(* Logix 5000 project; controller R400_500_XLS vendor 1 type 14 code 216 rev 31.11; software revision 31.01; part 32 of 32 *)
(* tags used below, declared in another part *)
   CycExcBuffer : UDT_CYCLE;
   CycleSequence : UDT_CYCLE_SEQUENCE;
   DRYING : DINT;   // Drying id number
   FINALRINSE_1 : DINT;   // Final rinse 1 id number
   M : DINT[5];   // Memory Bits
   OneShot : DINT[1];
   RINSE_4 : DINT;   // Rinse 4 id number
   RinseExcBuffer : UDT_RINSE;
   VENTING : DINT;   // Venting id number
   TreatmentPtr : DINT;
   Unit : Hrdwre;   // Unit Configuration
(* MainProgram, continued *)

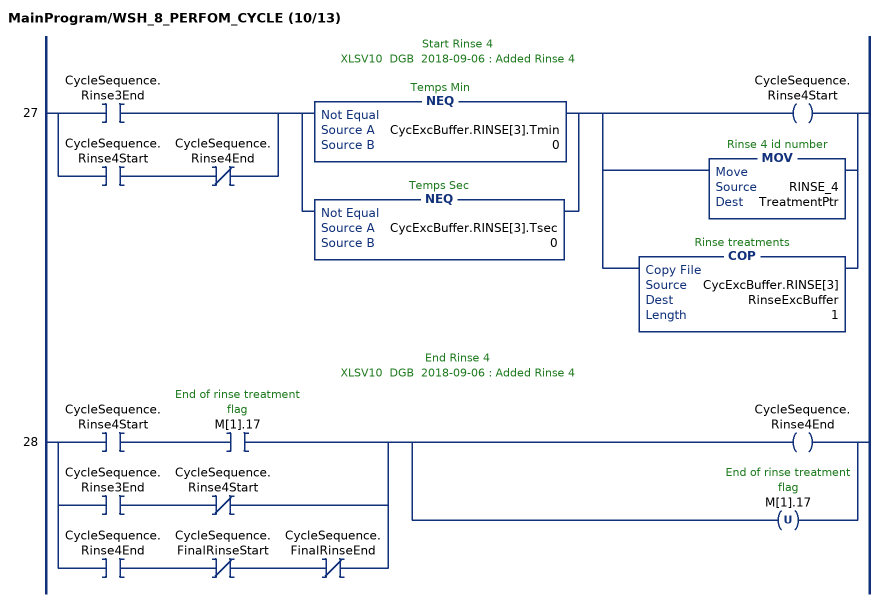
   [picture p660: MainProgram/WSH_8_PERFOM_CYCLE rungs 27-28]
   // Start Rinse 4
   // XLSV10  DGB  2018-09-06 : Added Rinse 4
   27: [XIC(CycleSequence.Rinse3End) ,XIC(CycleSequence.Rinse4Start) XIO(CycleSequence.Rinse4End) ][NEQ(CycExcBuffer.RINSE[3].Tmin,0) ,NEQ(CycExcBuffer.RINSE[3].Tsec,0) ][OTE(CycleSequence.Rinse4Start) ,MOV(RINSE_4,TreatmentPtr) ,COP(CycExcBuffer.RINSE[3],RinseExcBuffer,1) ];
   // End Rinse 4
   // XLSV10  DGB  2018-09-06 : Added Rinse 4
   28: [XIC(CycleSequence.Rinse4Start) XIC(M[1].17) ,XIC(CycleSequence.Rinse3End) XIO(CycleSequence.Rinse4Start) ,XIC(CycleSequence.Rinse4End) XIO(CycleSequence.FinalRinseStart) XIO(CycleSequence.FinalRinseEnd) ][OTE(CycleSequence.Rinse4End) ,OTU(M[1].17) ];
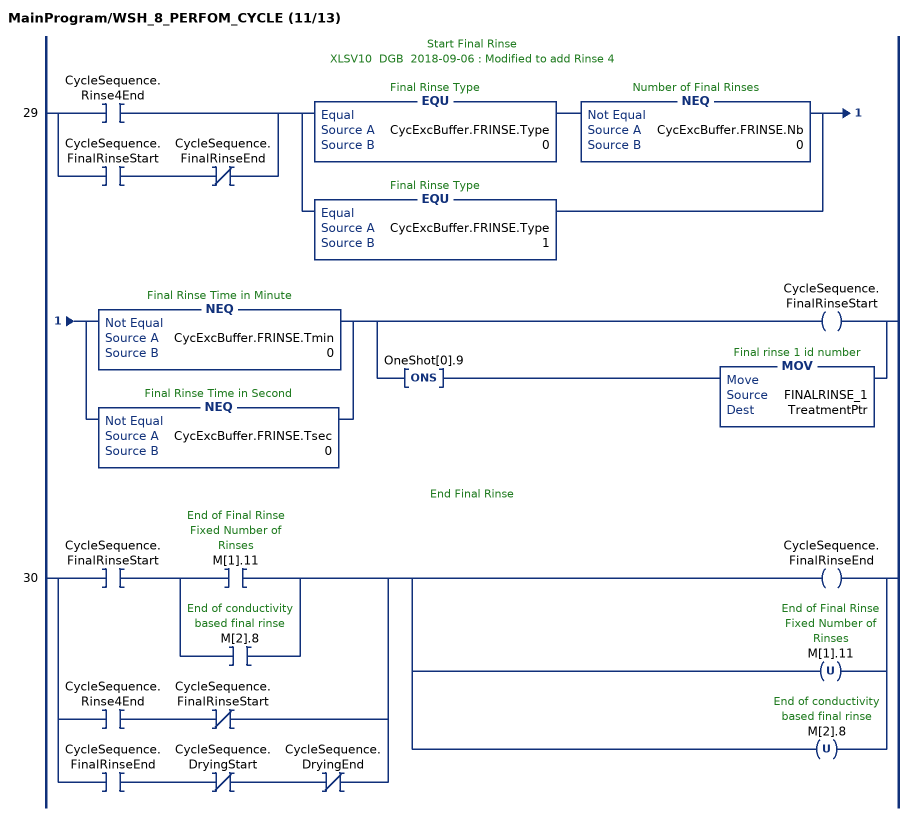
   // Start Final Rinse
   // XLSV10  DGB  2018-09-06 : Modified to add Rinse 4
   29: [XIC(CycleSequence.Rinse4End) ,XIC(CycleSequence.FinalRinseStart) XIO(CycleSequence.FinalRinseEnd) ][EQU(CycExcBuffer.FRINSE.Type,0) NEQ(CycExcBuffer.FRINSE.Nb,0) ,EQU(CycExcBuffer.FRINSE.Type,1) ][NEQ(CycExcBuffer.FRINSE.Tmin,0) ,NEQ(CycExcBuffer.FRINSE.Tsec,0) ][OTE(CycleSequence.FinalRinseStart) ,ONS(OneShot[0].9) MOV(FINALRINSE_1,TreatmentPtr) ];
   // End Final Rinse
   30: [XIC(CycleSequence.FinalRinseStart) [XIC(M[1].11) ,XIC(M[2].8) ] ,XIC(CycleSequence.Rinse4End) XIO(CycleSequence.FinalRinseStart) ,XIC(CycleSequence.FinalRinseEnd) XIO(CycleSequence.DryingStart) XIO(CycleSequence.DryingEnd) ][OTE(CycleSequence.FinalRinseEnd) ,OTU(M[1].11) ,OTU(M[2].8) ];
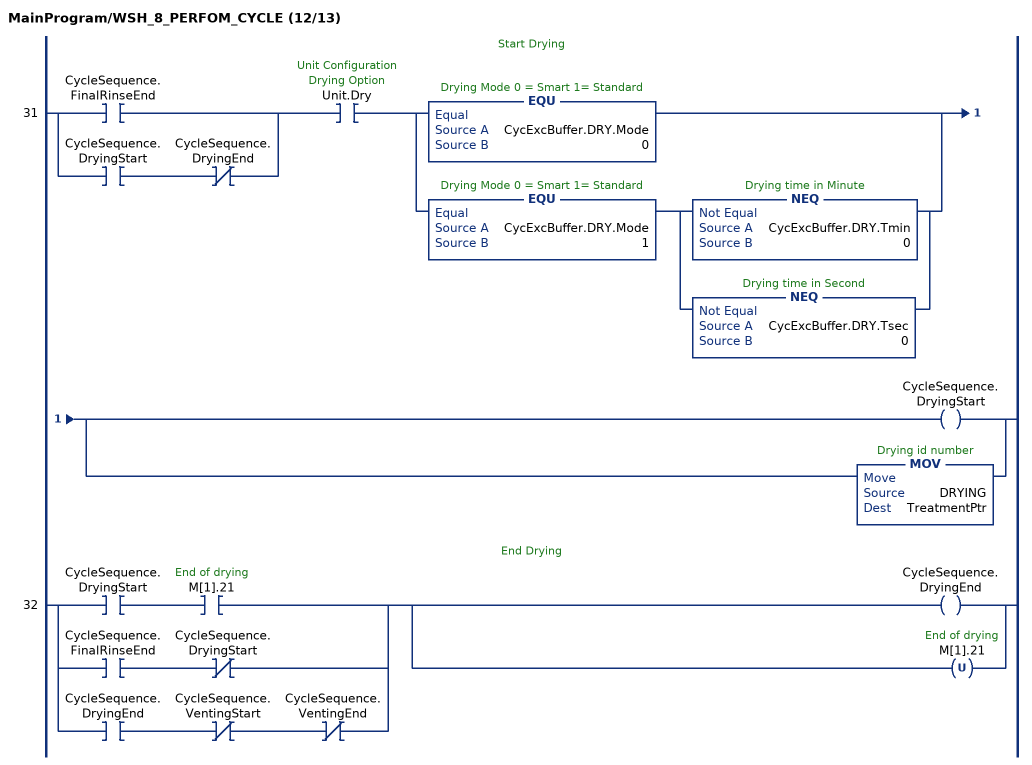
   // Start Drying
   31: [XIC(CycleSequence.FinalRinseEnd) ,XIC(CycleSequence.DryingStart) XIO(CycleSequence.DryingEnd) ]XIC(Unit.Dry)[EQU(CycExcBuffer.DRY.Mode,0) ,EQU(CycExcBuffer.DRY.Mode,1) [NEQ(CycExcBuffer.DRY.Tmin,0) ,NEQ(CycExcBuffer.DRY.Tsec,0) ] ][OTE(CycleSequence.DryingStart) ,MOV(DRYING,TreatmentPtr) ];
   // End Drying
   32: [XIC(CycleSequence.DryingStart) XIC(M[1].21) ,XIC(CycleSequence.FinalRinseEnd) XIO(CycleSequence.DryingStart) ,XIC(CycleSequence.DryingEnd) XIO(CycleSequence.VentingStart) XIO(CycleSequence.VentingEnd) ][OTE(CycleSequence.DryingEnd) ,OTU(M[1].21) ];
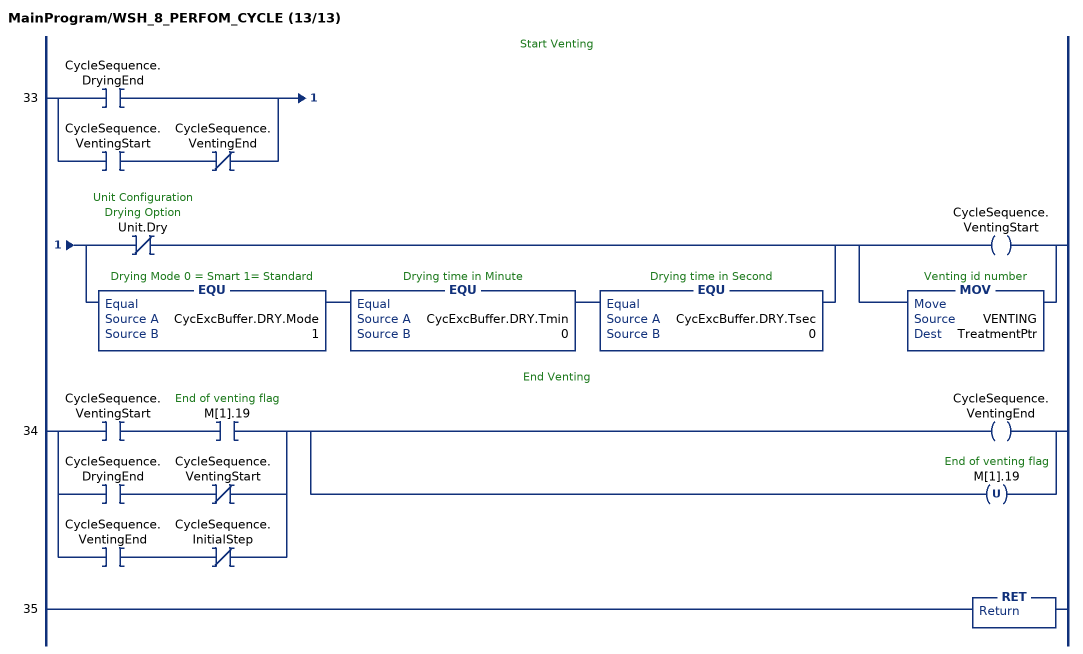
   // Start Venting
   33: [XIC(CycleSequence.DryingEnd) ,XIC(CycleSequence.VentingStart) XIO(CycleSequence.VentingEnd) ][XIO(Unit.Dry) ,EQU(CycExcBuffer.DRY.Mode,1) EQU(CycExcBuffer.DRY.Tmin,0) EQU(CycExcBuffer.DRY.Tsec,0) ][OTE(CycleSequence.VentingStart) ,MOV(VENTING,TreatmentPtr) ];
   // End Venting
   34: [XIC(CycleSequence.VentingStart) XIC(M[1].19) ,XIC(CycleSequence.DryingEnd) XIO(CycleSequence.VentingStart) ,XIC(CycleSequence.VentingEnd) XIO(CycleSequence.InitialStep) ][OTE(CycleSequence.VentingEnd) ,OTU(M[1].19) ];
   35: RET();
END_ROUTINE
END_PROGRAM
